// TIA Portal V20 export
// export: Created 2026-10-12T16:46:22.7550069Z, ExportSetting WithDefaults, DisplayName Totally Integrated Automation Portal, DisplayVersion V20 Update 6, DisplayName TIA Portal Openness, DisplayVersion V20 Update 6, DisplayName TIA Portal Version Control Interface, DisplayVersion V20 Update 6, DisplayName SINAMICS Startdrive Advanced, DisplayVersion V20 SP1 Update 2, DisplayName SINAMICS Startdrive G110M, G120, G120C, G120D, G120P, G115D, DisplayVersion V20 SP1 Update 2, DisplayName SINAMICS Startdrive G130, G150, S120, S150, SINAMICS MV, G220, S200, S210, DisplayVersion V20 SP1 Update 2, DisplayName STEP 7 Professional, DisplayVersion V20 Update 6, DisplayName STEP 7 Safety, DisplayVersion V20 Update 2, DisplayName WinCC Basic/Comfort/Advanced, DisplayVersion V20 Update 6, DisplayName WinCC Professional, DisplayVersion V20 Update 6, DisplayName WinCC Unified, DisplayVersion V20 Update 6
TYPE "UDT_FlexKraft_Device"
// ==============================================================================
//  UDT 3: Komplettes GerÃ¤t (Out + In zusammen, 64 Byte)
// ==============================================================================
// stored: IsFailsafeCompliant false
   STRUCT
      Out { S7_SetPoint := 'True'} : "UDT_FlexKraft_Out";   // 32 Byte SPS -> FK
      In { S7_SetPoint := 'True'} : "UDT_FlexKraft_In";   // 32 Byte FK -> SPS
   END_STRUCT;
END_TYPE
